(* IEC 61131-3 sources: kns-port-domestic/tools/plcopen/tests/fixtures/constructs/src/GVLs, 3 files *)

(* ---- GVL_Const.gvl.st ---- *)
// Константы
{attribute 'qualified_only'}
VAR_GLOBAL CONSTANT
    MAX_ITEMS : INT := 4;           // число элементов
    RATE_LIMIT : REAL := 0.25;
    TEXT_OK : STRING := 'OK';
END_VAR

(* ---- GVL_Io.gvl.st ---- *)
// Входы-выходы и сохраняемые значения
VAR_GLOBAL
    xDiStart AT %IX0.0 : BOOL;      // кнопка «Пуск»
    xDoRun AT %QX0.0 : BOOL;
    iAiLevel AT %IW2 : INT;
    astCmd : ARRAY[1..GVL_Const.MAX_ITEMS] OF ST_MotorCmd;
END_VAR
VAR_GLOBAL RETAIN
    udiRunHours : UDINT;
END_VAR
VAR_GLOBAL CONSTANT
    IO_CHANNELS : INT := 2;         // число каналов (константа в одном списке с переменными)
END_VAR

(* ---- PersistentVars.pvl.st ---- *)
// Сохраняемые переменные (объект Persistent Variables)
VAR_GLOBAL PERSISTENT RETAIN
    udiStartsTotal : UDINT;     // пуски за весь срок службы
    rRunHours_h : REAL;
END_VAR
